FUNCTION_BLOCK EmptyControl (* Extracted Composite Function Block Type *)
  (* Standard: 61499-2 *)
  (* Version 10/20/2026, lizar *)
  PACKAGE Main;
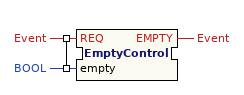
  EVENT_INPUT
    REQ WITH empty; (* Normal Execution Request *)
  END_EVENT
  EVENT_OUTPUT
    EMPTY;
  END_EVENT
  VAR_INPUT
    empty : BOOL;
  END_VAR
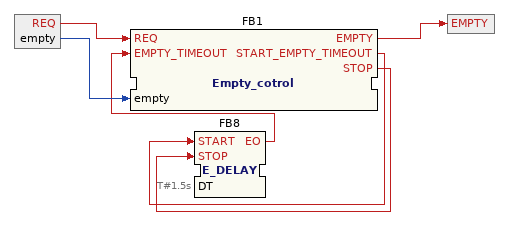
  FBS
    FB8 : E_DELAY(DT := T#1.5s);
    FB1 : Empty_cotrol;
  END_FBS
  EVENT_CONNECTIONS
    FB8.EO TO FB1.EMPTY_TIMEOUT;
    FB1.START_EMPTY_TIMEOUT TO FB8.START;
    FB1.STOP TO FB8.STOP;
    REQ TO FB1.REQ;
    FB1.EMPTY TO EMPTY;
  END_CONNECTIONS
  DATA_CONNECTIONS
    empty TO FB1.empty;
  END_CONNECTIONS
END_FUNCTION_BLOCK
